// TIA Portal V19 export
DATA_BLOCK "Tacho2_EM02"   // DB3
VERSION : 1.0
// stored: InstanceOfName EM02_Vacio, InstanceOfType FB
"EM02_Vacio"
   // VAR_INPUT
   //    In : "EM02_Input";
   //    VacuumPV : Real := 1000.0;
   //    PumpFbkRun : Bool;
   // END_VAR
   // VAR_OUTPUT
   //    Out : "EM02_Output";
   //    CM_PIC_MV : Real := 100.0;
   //    CM_MotL_Out : Bool := FALSE;
   //    CM_Bk_Out : Bool := FALSE;
   //    TimeoutAlarm : Bool := FALSE;
   //    SensorAlarm : Bool := FALSE;
   //    CMAlarm : Bool := FALSE;
   // END_VAR
   // VAR
   //    State : Int := 1;
   //    ActiveAction : Int := 1;
   //    AlarmLatched : Bool := TRUE;
   //    FaultCode : Int := 4;
   //    TimerReachedSP { S7_SetPoint := 'True'} : TON_TIME;
   //    TimerTimeout { S7_SetPoint := 'True'} : TON_TIME;
   //    TrigStart { S7_SetPoint := 'True'} : R_TRIG;
   //    TrigStop { S7_SetPoint := 'True'} : R_TRIG;
   //    TrigHold { S7_SetPoint := 'True'} : R_TRIG;
   //    TrigAbort { S7_SetPoint := 'True'} : R_TRIG;
   //    TrigReset { S7_SetPoint := 'True'} : R_TRIG;
   //    CM_PIC_Vacuum { S7_SetPoint := 'True'} : "PidL";
   //    CM_MotL { S7_SetPoint := 'True'} : "MotL";
   //    CM_Vlv_Break { S7_SetPoint := 'True'} : "VlvL";
   // END_VAR
BEGIN
   In.Cmds.Start := FALSE;
   In.Cmds.Stop := FALSE;
   In.Cmds.Hold := FALSE;
   In.Cmds.Abort := FALSE;
   In.Cmds.Reset := FALSE;
   In.Cmds.Manual := FALSE;
   In.Cmds.Auto := FALSE;
   In.Cmds.Maintenance := FALSE;
   In.CtrlMode := 0;
   In.VaccumSP := 200.0;
   In.AtmPressure := 980.0;
   In.VaccumValid := TRUE;
   In.VaccumFilter := T#3S;
   In.VaccumTimeout := T#10M;
   In.VaccumSMMV := 0.0;
   Out.Status.ModeMan := FALSE;
   Out.Status.ModeAuto := TRUE;
   Out.Status.ModeMaint := FALSE;
   Out.Status.ModeConflict := FALSE;
   Out.Status.Idle := FALSE;
   Out.Status.Running := TRUE;
   Out.Status.Completed := FALSE;
   Out.Status.Holding := FALSE;
   Out.Status.Held := FALSE;
   Out.Status.Stopping := FALSE;
   Out.Status.Stopped := FALSE;
   Out.Status.Aborting := FALSE;
   Out.Status.Aborted := FALSE;
   Out.Status.Fault := TRUE;
   Out.Status.State := 1;
   Out.Status.FaultCode := 4;
   Out.VacuumActive := TRUE;
   Out.VacuumBroken := FALSE;
   TimerReachedSP.PT := T#0MS;
   TimerReachedSP.IN := FALSE;
   TimerTimeout.PT := T#10M;
   TimerTimeout.IN := TRUE;
   TrigStart.CLK := TRUE;
   TrigStart.Q := FALSE;
   TrigStart.Stat_Bit := TRUE;
   TrigStop.CLK := FALSE;
   TrigStop.Q := FALSE;
   TrigStop.Stat_Bit := FALSE;
   TrigHold.CLK := FALSE;
   TrigHold.Q := FALSE;
   TrigHold.Stat_Bit := FALSE;
   TrigAbort.CLK := FALSE;
   TrigAbort.Q := FALSE;
   TrigAbort.Stat_Bit := FALSE;
   TrigReset.CLK := FALSE;
   TrigReset.Q := FALSE;
   TrigReset.Stat_Bit := FALSE;
   CM_PIC_Vacuum.AutModLi := TRUE;
   CM_PIC_Vacuum.ManModLi := FALSE;
   CM_PIC_Vacuum.LocModLi := FALSE;
   CM_PIC_Vacuum.OosModLi := FALSE;
   CM_PIC_Vacuum.ModLiOp := TRUE;
   CM_PIC_Vacuum.ResetLi := FALSE;
   CM_PIC_Vacuum.SPModLiOp := TRUE;
   CM_PIC_Vacuum.ExtModLi := FALSE;
   CM_PIC_Vacuum.IntModLi := TRUE;
   CM_PIC_Vacuum.PV := 1000.0;
   CM_PIC_Vacuum.PV_Norm.High := 2000.0;
   CM_PIC_Vacuum.PV_Norm.Low := 0.0;
   CM_PIC_Vacuum.MV_Norm.High := 100.0;
   CM_PIC_Vacuum.MV_Norm.Low := 0.0;
   CM_PIC_Vacuum.PV_Scale.High := 2000.0;
   CM_PIC_Vacuum.PV_Scale.Low := 0.0;
   CM_PIC_Vacuum.SPExt := 0.0;
   CM_PIC_Vacuum.SP_HiLim := 2000.0;
   CM_PIC_Vacuum.SP_LoLim := 0.0;
   CM_PIC_Vacuum.MV_HiLim := 100.0;
   CM_PIC_Vacuum.MV_LoLim := 0.0;
   CM_PIC_Vacuum.OosSafeMV := 0.0;
   CM_PIC_Vacuum.PV_unit := 1138;
   CM_PIC_Vacuum.MV_unit := 1342;
   CM_PIC_Vacuum.DataHMI.identName := 'PCV-210';
   CM_PIC_Vacuum.DataHMI.comment := 'Vacio';
   CM_PIC_Vacuum.DataHMI.AutModOp := TRUE;
   CM_PIC_Vacuum.DataHMI.ManModOp := FALSE;
   CM_PIC_Vacuum.DataHMI.LocModOp := FALSE;
   CM_PIC_Vacuum.DataHMI.OosModOp := FALSE;
   CM_PIC_Vacuum.DataHMI.ResetOp := FALSE;
   CM_PIC_Vacuum.DataHMI.MonitorOn := FALSE;
   CM_PIC_Vacuum.DataHMI.ExtModOp := FALSE;
   CM_PIC_Vacuum.DataHMI.IntModOp := FALSE;
   CM_PIC_Vacuum.DataHMI.SpInt := 200.0;
   CM_PIC_Vacuum.DataHMI.Man := 100.0;
   CM_PIC_Vacuum.DataHMI.PermissionLog.AutModOpEn := FALSE;
   CM_PIC_Vacuum.DataHMI.PermissionLog.ManModOpEn := FALSE;
   CM_PIC_Vacuum.DataHMI.PermissionLog.LocModOpEn := FALSE;
   CM_PIC_Vacuum.DataHMI.PermissionLog.OosModOpEn := FALSE;
   CM_PIC_Vacuum.DataHMI.PermissionLog.ResetOpEn := TRUE;
   CM_PIC_Vacuum.DataHMI.PermissionLog.ExtModOpEn := FALSE;
   CM_PIC_Vacuum.DataHMI.PermissionLog.IntModOpEn := FALSE;
   CM_PIC_Vacuum.DataHMI.PermissionLog.Alarms.MsgSupEn := FALSE;
   CM_PIC_Vacuum.DataHMI.PermissionLog.Alarms.HiAlmSupEn := FALSE;
   CM_PIC_Vacuum.DataHMI.PermissionLog.Alarms.HiWrnSupEn := FALSE;
   CM_PIC_Vacuum.DataHMI.PermissionLog.Alarms.LoWrnSupEn := FALSE;
   CM_PIC_Vacuum.DataHMI.PermissionLog.Alarms.LoAlmSupEn := FALSE;
   CM_PIC_Vacuum.DataHMI.Status.OosAct := FALSE;
   CM_PIC_Vacuum.DataHMI.Status.LocAct := FALSE;
   CM_PIC_Vacuum.DataHMI.Status.ManAct := FALSE;
   CM_PIC_Vacuum.DataHMI.Status.AutAct := TRUE;
   CM_PIC_Vacuum.DataHMI.Status.SpExtAct := FALSE;
   CM_PIC_Vacuum.DataHMI.Status.Protection := FALSE;
   CM_PIC_Vacuum.DataHMI.Status.Intlock := TRUE;
   CM_PIC_Vacuum.DataHMI.Status.Permit := TRUE;
   CM_PIC_Vacuum.DataHMI.Status.TrackAct := FALSE;
   CM_PIC_Vacuum.DataHMI.Status.SP := 200.0;
   CM_PIC_Vacuum.DataHMI.Status.PV := 1000.0;
   CM_PIC_Vacuum.DataHMI.Status.ER := -800.0;
   CM_PIC_Vacuum.DataHMI.Status.MV := 100.0;
   CM_PIC_Vacuum.DataHMI.Status.PVOpScale.High := 2000.0;
   CM_PIC_Vacuum.DataHMI.Status.PVOpScale.Low := 0.0;
   CM_PIC_Vacuum.DataHMI.Status.MVOpScale.High := 100.0;
   CM_PIC_Vacuum.DataHMI.Status.MVOpScale.Low := 0.0;
   CM_PIC_Vacuum.DataHMI.Status.SPIntLim.High := 0.0;
   CM_PIC_Vacuum.DataHMI.Status.SPIntLim.Low := 0.0;
   CM_PIC_Vacuum.DataHMI.Status.PV_unit := 1138;
   CM_PIC_Vacuum.DataHMI.Status.MV_unit := 1342;
   CM_PIC_Vacuum.DataHMI.PIDConfig.NegGain := TRUE;
   CM_PIC_Vacuum.DataHMI.PIDConfig.P_Sel := TRUE;
   CM_PIC_Vacuum.DataHMI.PIDConfig.I_Sel := TRUE;
   CM_PIC_Vacuum.DataHMI.PIDConfig.D_Sel := FALSE;
   CM_PIC_Vacuum.DataHMI.PIDConfig.Gain := -2.0;
   CM_PIC_Vacuum.DataHMI.PIDConfig.Ti := 20.0;
   CM_PIC_Vacuum.DataHMI.PIDConfig.Td := 10.0;
   CM_PIC_Vacuum.DataHMI.PIDConfig.DeadBW := 0.0;
   CM_PIC_Vacuum.DataHMI.Alarms.identName := 'PCV-210';
   CM_PIC_Vacuum.DataHMI.Alarms.comment := 'Vacio';
   CM_PIC_Vacuum.DataHMI.Alarms.MsgSupOp := FALSE;
   CM_PIC_Vacuum.DataHMI.Alarms.PVScale.High := 2000.0;
   CM_PIC_Vacuum.DataHMI.Alarms.PVScale.Low := 0.0;
   CM_PIC_Vacuum.DataHMI.Alarms.HiAlmSupOp := FALSE;
   CM_PIC_Vacuum.DataHMI.Alarms.HiWrnSupOp := FALSE;
   CM_PIC_Vacuum.DataHMI.Alarms.LoWrnSupOp := FALSE;
   CM_PIC_Vacuum.DataHMI.Alarms.LoAlmSupOp := FALSE;
   CM_PIC_Vacuum.DataHMI.Alarms.PermissionLog.MsgSupEn := FALSE;
   CM_PIC_Vacuum.DataHMI.Alarms.PermissionLog.HiAlmSupEn := TRUE;
   CM_PIC_Vacuum.DataHMI.Alarms.PermissionLog.HiWrnSupEn := TRUE;
   CM_PIC_Vacuum.DataHMI.Alarms.PermissionLog.LoWrnSupEn := TRUE;
   CM_PIC_Vacuum.DataHMI.Alarms.PermissionLog.LoAlmSupEn := TRUE;
   CM_PIC_Vacuum.DataHMI.Alarms.Status.PV := 1000.0;
   CM_PIC_Vacuum.DataHMI.Alarms.Status.PV_unit := 1138;
   CM_PIC_Vacuum.DataHMI.Alarms.Status.PV_HiAlm := TRUE;
   CM_PIC_Vacuum.DataHMI.Alarms.Status.PV_HiWrn := TRUE;
   CM_PIC_Vacuum.DataHMI.Alarms.Status.PV_LoWrn := FALSE;
   CM_PIC_Vacuum.DataHMI.Alarms.Status.PV_LoAlm := FALSE;
   CM_PIC_Vacuum.DataHMI.Alarms.Status.MsgSup := FALSE;
   CM_PIC_Vacuum.Feature.Startup := TRUE;
   CM_PIC_Vacuum.Feature.MSSOff := TRUE;
   CM_PIC_Vacuum.Feature.FltOff := TRUE;
   CM_PIC_Vacuum.Feature.LocalMod := FALSE;
   CM_PIC_Vacuum.Permission.AutModOpEn := TRUE;
   CM_PIC_Vacuum.Permission.ManModOpEn := TRUE;
   CM_PIC_Vacuum.Permission.LocModOpEn := FALSE;
   CM_PIC_Vacuum.Permission.OosModOpEn := FALSE;
   CM_PIC_Vacuum.Permission.ResetOpEn := TRUE;
   CM_PIC_Vacuum.Permission.ExtModOpEn := FALSE;
   CM_PIC_Vacuum.Permission.IntModOpEn := TRUE;
   CM_PIC_Vacuum.Permission.Alarms.MsgSupEn := TRUE;
   CM_PIC_Vacuum.Permission.Alarms.HiAlmSupEn := TRUE;
   CM_PIC_Vacuum.Permission.Alarms.HiWrnSupEn := TRUE;
   CM_PIC_Vacuum.Permission.Alarms.LoWrnSupEn := TRUE;
   CM_PIC_Vacuum.Permission.Alarms.LoAlmSupEn := TRUE;
   CM_PIC_Vacuum.MSS := TRUE;
   CM_PIC_Vacuum.Trip := FALSE;
   CM_PIC_Vacuum.Permit := TRUE;
   CM_PIC_Vacuum.Intlock := TRUE;
   CM_PIC_Vacuum.Protect := TRUE;
   CM_PIC_Vacuum.TrackOn := FALSE;
   CM_PIC_Vacuum.Rbk := 0.0;
   CM_PIC_Vacuum.RbkHiTol := 3.0;
   CM_PIC_Vacuum.RbkLoTol := 3.0;
   CM_PIC_Vacuum.RbkMonTime := T#3S;
   CM_PIC_Vacuum.TrackVal := 0.0;
   CM_PIC_Vacuum.RunUpCyc := 3;
   CM_PIC_Vacuum.DisV := 0.0;
   CM_PIC_Vacuum.HiAlm := 95.0;
   CM_PIC_Vacuum.HiWrn := 90.0;
   CM_PIC_Vacuum.LoWrn := 10.0;
   CM_PIC_Vacuum.LoAlm := 5.0;
   CM_PIC_Vacuum.Hyst := 5.0;
   CM_PIC_Vacuum.AutAct := TRUE;
   CM_PIC_Vacuum.ManAct := FALSE;
   CM_PIC_Vacuum.LocAct := FALSE;
   CM_PIC_Vacuum.OosAct := FALSE;
   CM_PIC_Vacuum.MsgSup := TRUE;
   CM_PIC_Vacuum.AlarmError := FALSE;
   CM_PIC_Vacuum.MV := 100.0;
   CM_PIC_Vacuum.SPExtAct := FALSE;
   CM_PIC_Vacuum.SP := 200.0;
   CM_PIC_Vacuum.ER := -800.0;
   CM_PIC_Vacuum.PVH_Alm := TRUE;
   CM_PIC_Vacuum.PVH_Wrn := TRUE;
   CM_PIC_Vacuum.PVL_Wrn := FALSE;
   CM_PIC_Vacuum.PVL_Alm := FALSE;
   CM_PIC_Vacuum.controller.COM_RST := FALSE;
   CM_PIC_Vacuum.controller.MAN_ON := FALSE;
   CM_PIC_Vacuum.controller.PVPER_ON := FALSE;
   CM_PIC_Vacuum.controller.P_SEL := TRUE;
   CM_PIC_Vacuum.controller.I_SEL := TRUE;
   CM_PIC_Vacuum.controller.INT_HOLD := FALSE;
   CM_PIC_Vacuum.controller.I_ITL_ON := FALSE;
   CM_PIC_Vacuum.controller.D_SEL := FALSE;
   CM_PIC_Vacuum.controller.CYCLE := T#1S;
   CM_PIC_Vacuum.controller.SP_INT := 10.0;
   CM_PIC_Vacuum.controller.PV_IN := 50.0;
   CM_PIC_Vacuum.controller.PV_PER := 16#0000;
   CM_PIC_Vacuum.controller.MAN := 100.0;
   CM_PIC_Vacuum.controller.GAIN := -2.0;
   CM_PIC_Vacuum.controller.TI := T#20S;
   CM_PIC_Vacuum.controller.TD := T#10S;
   CM_PIC_Vacuum.controller.TM_LAG := T#2S;
   CM_PIC_Vacuum.controller.DEADB_W := 0.0;
   CM_PIC_Vacuum.controller.LMN_HLM := 100.0;
   CM_PIC_Vacuum.controller.LMN_LLM := 0.0;
   CM_PIC_Vacuum.controller.PV_FAC := 1.0;
   CM_PIC_Vacuum.controller.PV_OFF := 0.0;
   CM_PIC_Vacuum.controller.LMN_FAC := 1.0;
   CM_PIC_Vacuum.controller.LMN_OFF := 0.0;
   CM_PIC_Vacuum.controller.I_ITLVAL := 0.0;
   CM_PIC_Vacuum.controller.DISV := 0.0;
   CM_PIC_Vacuum.controller.LMN := 100.0;
   CM_PIC_Vacuum.controller.LMN_PER := 16#6C00;
   CM_PIC_Vacuum.controller.QLMN_HLM := TRUE;
   CM_PIC_Vacuum.controller.QLMN_LLM := FALSE;
   CM_PIC_Vacuum.controller.LMN_P := 80.0;
   CM_PIC_Vacuum.controller.LMN_I := 80.0;
   CM_PIC_Vacuum.controller.LMN_D := 0.0;
   CM_PIC_Vacuum.controller.PV := 50.0;
   CM_PIC_Vacuum.controller.ER := -40.0;
   CM_PIC_Vacuum.controller.sInvAlt := 80.0;
   CM_PIC_Vacuum.controller.sIanteilAlt := 80.0;
   CM_PIC_Vacuum.controller.sRestInt := 0.0;
   CM_PIC_Vacuum.controller.sRestDif := 0.0;
   CM_PIC_Vacuum.controller.sRueck := 80.0;
   CM_PIC_Vacuum.controller.sLmn := 100.0;
   CM_PIC_Vacuum.controller.sbArwHLmOn := TRUE;
   CM_PIC_Vacuum.controller.sbArwLLmOn := FALSE;
   CM_PIC_Vacuum.controller.sbILimOn := TRUE;
   CM_PIC_Vacuum.ModSelInt := 2;
   CM_PIC_Vacuum.stRestart := FALSE;
   CM_PIC_Vacuum.ResetLiLogic := FALSE;
   CM_PIC_Vacuum.ResetResult := FALSE;
   CM_PIC_Vacuum.stResetLiLogic := FALSE;
   CM_PIC_Vacuum.stMonErr := FALSE;
   CM_PIC_Vacuum.stTripErr := FALSE;
   CM_PIC_Vacuum.stProtErr := FALSE;
   CM_PIC_Vacuum.stMSS := FALSE;
   CM_PIC_Vacuum.stProt := FALSE;
   CM_PIC_Vacuum.stTrip := FALSE;
   CM_PIC_Vacuum.stLockFault := FALSE;
   CM_PIC_Vacuum.stRun := FALSE;
   CM_PIC_Vacuum.stExtMod := FALSE;
   CM_PIC_Vacuum.stAutoLogic := FALSE;
   CM_PIC_Vacuum.RuntimeMem := 16#0000_0EAA_9B49_C0F5;
   CM_PIC_Vacuum.RuntimeS := 0.999710415986597;
   CM_PIC_Vacuum.PVMon.Feature.Startup := TRUE;
   CM_PIC_Vacuum.PVMon.Enable := TRUE;
   CM_PIC_Vacuum.PVMon.Permission.MsgSupEn := TRUE;
   CM_PIC_Vacuum.PVMon.Permission.HiAlmSupEn := TRUE;
   CM_PIC_Vacuum.PVMon.Permission.HiWrnSupEn := TRUE;
   CM_PIC_Vacuum.PVMon.Permission.LoWrnSupEn := TRUE;
   CM_PIC_Vacuum.PVMon.Permission.LoAlmSupEn := TRUE;
   CM_PIC_Vacuum.PVMon.DataHMI.identName := 'PCV-210';
   CM_PIC_Vacuum.PVMon.DataHMI.comment := 'Vacio';
   CM_PIC_Vacuum.PVMon.DataHMI.MsgSupOp := FALSE;
   CM_PIC_Vacuum.PVMon.DataHMI.PVScale.High := 2000.0;
   CM_PIC_Vacuum.PVMon.DataHMI.PVScale.Low := 0.0;
   CM_PIC_Vacuum.PVMon.DataHMI.HiAlmSupOp := FALSE;
   CM_PIC_Vacuum.PVMon.DataHMI.HiWrnSupOp := FALSE;
   CM_PIC_Vacuum.PVMon.DataHMI.LoWrnSupOp := FALSE;
   CM_PIC_Vacuum.PVMon.DataHMI.LoAlmSupOp := FALSE;
   CM_PIC_Vacuum.PVMon.DataHMI.PermissionLog.MsgSupEn := FALSE;
   CM_PIC_Vacuum.PVMon.DataHMI.PermissionLog.HiAlmSupEn := TRUE;
   CM_PIC_Vacuum.PVMon.DataHMI.PermissionLog.HiWrnSupEn := TRUE;
   CM_PIC_Vacuum.PVMon.DataHMI.PermissionLog.LoWrnSupEn := TRUE;
   CM_PIC_Vacuum.PVMon.DataHMI.PermissionLog.LoAlmSupEn := TRUE;
   CM_PIC_Vacuum.PVMon.DataHMI.Status.PV := 1000.0;
   CM_PIC_Vacuum.PVMon.DataHMI.Status.PV_unit := 1138;
   CM_PIC_Vacuum.PVMon.DataHMI.Status.PV_HiAlm := TRUE;
   CM_PIC_Vacuum.PVMon.DataHMI.Status.PV_HiWrn := TRUE;
   CM_PIC_Vacuum.PVMon.DataHMI.Status.PV_LoWrn := FALSE;
   CM_PIC_Vacuum.PVMon.DataHMI.Status.PV_LoAlm := FALSE;
   CM_PIC_Vacuum.PVMon.DataHMI.Status.MsgSup := FALSE;
   CM_PIC_Vacuum.PVMon.RunUpCyc := 3;
   CM_PIC_Vacuum.PVMon.PV := 1000.0;
   CM_PIC_Vacuum.PVMon.HiAlm := 95.0;
   CM_PIC_Vacuum.PVMon.HiWrn := 90.0;
   CM_PIC_Vacuum.PVMon.LoWrn := 10.0;
   CM_PIC_Vacuum.PVMon.LoAlm := 5.0;
   CM_PIC_Vacuum.PVMon.Hyst := 5.0;
   CM_PIC_Vacuum.PVMon.PV_unit := 1138;
   CM_PIC_Vacuum.PVMon.MsgErr := FALSE;
   CM_PIC_Vacuum.PVMon.MsgSup := TRUE;
   CM_PIC_Vacuum.PVMon.PVH_Alm := TRUE;
   CM_PIC_Vacuum.PVMon.PVH_Wrn := TRUE;
   CM_PIC_Vacuum.PVMon.PVL_Wrn := FALSE;
   CM_PIC_Vacuum.PVMon.PVL_Alm := FALSE;
   CM_PIC_Vacuum.PVMon.stRestart := FALSE;
   CM_PIC_Vacuum.PVMon.RunUpCounter := 0;
   CM_PIC_Vacuum.PVMon.pSIG1 := TRUE;
   CM_PIC_Vacuum.PVMon.pSIG2 := TRUE;
   CM_PIC_Vacuum.PVMon.pSIG3 := FALSE;
   CM_PIC_Vacuum.PVMon.pSIG4 := FALSE;
   CM_PIC_Vacuum.PVMon.pAlarm := TRUE;
   CM_PIC_Vacuum.RunUpCounter := 0;
   CM_PIC_Vacuum.pAlarm := TRUE;
   CM_PIC_Vacuum.stMSSErr := FALSE;
   CM_PIC_Vacuum.SPMod := FALSE;
   CM_PIC_Vacuum.SPSelInt := 1;
   CM_PIC_Vacuum.stErr := FALSE;
   CM_PIC_Vacuum.stDivErr := FALSE;
   CM_PIC_Vacuum.stNegGain := TRUE;
   CM_PIC_Vacuum.stGain := -2.0;
   CM_PIC_Vacuum.stTi := 0.0;
   CM_PIC_Vacuum.stTd := 0.0;
   CM_PIC_Vacuum.stPIDConfig.NegGain := TRUE;
   CM_PIC_Vacuum.stPIDConfig.P_Sel := TRUE;
   CM_PIC_Vacuum.stPIDConfig.I_Sel := TRUE;
   CM_PIC_Vacuum.stPIDConfig.D_Sel := FALSE;
   CM_PIC_Vacuum.stPIDConfig.Gain := -2.0;
   CM_PIC_Vacuum.stPIDConfig.Ti := 20.0;
   CM_PIC_Vacuum.stPIDConfig.Td := 10.0;
   CM_PIC_Vacuum.stPIDConfig.DeadBW := 0.0;
   CM_PIC_Vacuum.RbkMonitorTimer.PT := T#0MS;
   CM_PIC_Vacuum.RbkMonitorTimer.IN := FALSE;
   CM_MotL.SampleT := 1.0;
   CM_MotL.AutModLi := TRUE;
   CM_MotL.ManModLi := FALSE;
   CM_MotL.LocModLi := FALSE;
   CM_MotL.OosModLi := FALSE;
   CM_MotL.ModLiOp := TRUE;
   CM_MotL.ResetLi := FALSE;
   CM_MotL.DataHMI.identName := 'M-102';
   CM_MotL.DataHMI.comment := 'Bba Vacio';
   CM_MotL.DataHMI.AutModOp := TRUE;
   CM_MotL.DataHMI.ManModOp := FALSE;
   CM_MotL.DataHMI.LocModOp := FALSE;
   CM_MotL.DataHMI.OosModOp := FALSE;
   CM_MotL.DataHMI.StartOp := FALSE;
   CM_MotL.DataHMI.StopOp := FALSE;
   CM_MotL.DataHMI.ResetOp := FALSE;
   CM_MotL.DataHMI.MonitorOn := FALSE;
   CM_MotL.DataHMI.PermissionLog.AutModOpEn := FALSE;
   CM_MotL.DataHMI.PermissionLog.ManModOpEn := FALSE;
   CM_MotL.DataHMI.PermissionLog.LocModOpEn := FALSE;
   CM_MotL.DataHMI.PermissionLog.OosModOpEn := FALSE;
   CM_MotL.DataHMI.PermissionLog.ResetOpEn := TRUE;
   CM_MotL.DataHMI.PermissionLog.StartOpEn := FALSE;
   CM_MotL.DataHMI.PermissionLog.StopOpEn := FALSE;
   CM_MotL.DataHMI.Status.OosAct := FALSE;
   CM_MotL.DataHMI.Status.LocAct := FALSE;
   CM_MotL.DataHMI.Status.ManAct := FALSE;
   CM_MotL.DataHMI.Status.AutAct := TRUE;
   CM_MotL.DataHMI.Status.CmdOnOff := TRUE;
   CM_MotL.DataHMI.Status.Run := TRUE;
   CM_MotL.DataHMI.Status.Stop := FALSE;
   CM_MotL.DataHMI.Status.MonErr := FALSE;
   CM_MotL.DataHMI.Status.Trip := FALSE;
   CM_MotL.DataHMI.Status.Protection := FALSE;
   CM_MotL.DataHMI.Status.Intlock := TRUE;
   CM_MotL.DataHMI.Status.Permit := TRUE;
   CM_MotL.DataHMI.MonitorTime := 3.0;
   CM_MotL.Feature.Startup := TRUE;
   CM_MotL.Feature.MSSOff := TRUE;
   CM_MotL.Feature.FltOff := TRUE;
   CM_MotL.Feature.LocalMod := FALSE;
   CM_MotL.Permission.AutModOpEn := TRUE;
   CM_MotL.Permission.ManModOpEn := TRUE;
   CM_MotL.Permission.LocModOpEn := FALSE;
   CM_MotL.Permission.OosModOpEn := FALSE;
   CM_MotL.Permission.ResetOpEn := TRUE;
   CM_MotL.Permission.StartOpEn := TRUE;
   CM_MotL.Permission.StopOpEn := TRUE;
   CM_MotL.MSS := TRUE;
   CM_MotL.Trip := FALSE;
   CM_MotL.Permit := TRUE;
   CM_MotL.Intlock := TRUE;
   CM_MotL.Protect := TRUE;
   CM_MotL.StartAut := TRUE;
   CM_MotL.StopAut := FALSE;
   CM_MotL.StartLoc := FALSE;
   CM_MotL.StopLoc := FALSE;
   CM_MotL.LockOn := FALSE;
   CM_MotL.FbkRun := FALSE;
   CM_MotL.RunUpCyc := 3;
   CM_MotL.Start := TRUE;
   CM_MotL.AutAct := TRUE;
   CM_MotL.ManAct := FALSE;
   CM_MotL.LocAct := FALSE;
   CM_MotL.OosAct := FALSE;
   CM_MotL.Run := TRUE;
   CM_MotL.Stop := FALSE;
   CM_MotL.MsgSup := FALSE;
   CM_MotL.AlarmError := FALSE;
   CM_MotL.ModSelInt := 2;
   CM_MotL.stRestart := FALSE;
   CM_MotL.ResetLiLogic := FALSE;
   CM_MotL.ResetResult := FALSE;
   CM_MotL.stResetLiLogic := FALSE;
   CM_MotL.stMonErr := FALSE;
   CM_MotL.stTripErr := FALSE;
   CM_MotL.stProtErr := FALSE;
   CM_MotL.stMSS := FALSE;
   CM_MotL.stProt := FALSE;
   CM_MotL.stTrip := FALSE;
   CM_MotL.stLockFault := FALSE;
   CM_MotL.stRun := TRUE;
   CM_MotL.stCmdOnOff := TRUE;
   CM_MotL.stAutoLogic := TRUE;
   CM_MotL.stbCmdOnOff := TRUE;
   CM_MotL.stActiveTime := 0.0;
   CM_MotL.RunUpCounter := 0;
   CM_MotL.pAlarm := TRUE;
   CM_MotL.stMSSErr := FALSE;
   CM_Vlv_Break.SampleT := 1.0;
   CM_Vlv_Break.AutModLi := TRUE;
   CM_Vlv_Break.ManModLi := FALSE;
   CM_Vlv_Break.LocModLi := FALSE;
   CM_Vlv_Break.OosModLi := FALSE;
   CM_Vlv_Break.ModLiOp := TRUE;
   CM_Vlv_Break.ResetLi := FALSE;
   CM_Vlv_Break.DataHMI.identName := 'PSV-103';
   CM_Vlv_Break.DataHMI.comment := 'Rompevacio';
   CM_Vlv_Break.DataHMI.AutModOp := TRUE;
   CM_Vlv_Break.DataHMI.ManModOp := FALSE;
   CM_Vlv_Break.DataHMI.LocModOp := FALSE;
   CM_Vlv_Break.DataHMI.OosModOp := FALSE;
   CM_Vlv_Break.DataHMI.OpenOp := FALSE;
   CM_Vlv_Break.DataHMI.CloseOp := FALSE;
   CM_Vlv_Break.DataHMI.ResetOp := FALSE;
   CM_Vlv_Break.DataHMI.MonitorOn := FALSE;
   CM_Vlv_Break.DataHMI.PermissionLog.AutModOpEn := FALSE;
   CM_Vlv_Break.DataHMI.PermissionLog.ManModOpEn := FALSE;
   CM_Vlv_Break.DataHMI.PermissionLog.LocModOpEn := FALSE;
   CM_Vlv_Break.DataHMI.PermissionLog.OosModOpEn := FALSE;
   CM_Vlv_Break.DataHMI.PermissionLog.ResetOpEn := TRUE;
   CM_Vlv_Break.DataHMI.PermissionLog.OpenOpEn := FALSE;
   CM_Vlv_Break.DataHMI.PermissionLog.CloseOpEn := FALSE;
   CM_Vlv_Break.DataHMI.Status.OosAct := FALSE;
   CM_Vlv_Break.DataHMI.Status.LocAct := FALSE;
   CM_Vlv_Break.DataHMI.Status.ManAct := FALSE;
   CM_Vlv_Break.DataHMI.Status.AutAct := TRUE;
   CM_Vlv_Break.DataHMI.Status.Cmd := FALSE;
   CM_Vlv_Break.DataHMI.Status.Opened := FALSE;
   CM_Vlv_Break.DataHMI.Status.Closed := TRUE;
   CM_Vlv_Break.DataHMI.Status.MonErr := FALSE;
   CM_Vlv_Break.DataHMI.Status.Trip := FALSE;
   CM_Vlv_Break.DataHMI.Status.Protection := FALSE;
   CM_Vlv_Break.DataHMI.Status.Intlock := FALSE;
   CM_Vlv_Break.DataHMI.Status.Permit := FALSE;
   CM_Vlv_Break.DataHMI.MonitorTime := 3.0;
   CM_Vlv_Break.Feature.Startup := TRUE;
   CM_Vlv_Break.Feature.MSSOff := TRUE;
   CM_Vlv_Break.Feature.FltOff := TRUE;
   CM_Vlv_Break.Feature.LocalMod := FALSE;
   CM_Vlv_Break.Permission.AutModOpEn := TRUE;
   CM_Vlv_Break.Permission.ManModOpEn := TRUE;
   CM_Vlv_Break.Permission.LocModOpEn := FALSE;
   CM_Vlv_Break.Permission.OosModOpEn := FALSE;
   CM_Vlv_Break.Permission.ResetOpEn := TRUE;
   CM_Vlv_Break.Permission.OpenOpEn := TRUE;
   CM_Vlv_Break.Permission.CloseOpEn := TRUE;
   CM_Vlv_Break.MSS := TRUE;
   CM_Vlv_Break.Trip := FALSE;
   CM_Vlv_Break.Permit := FALSE;
   CM_Vlv_Break.Intlock := FALSE;
   CM_Vlv_Break.Protect := TRUE;
   CM_Vlv_Break.OpenAut := FALSE;
   CM_Vlv_Break.CloseAut := TRUE;
   CM_Vlv_Break.OpenLoc := FALSE;
   CM_Vlv_Break.CloseLoc := FALSE;
   CM_Vlv_Break.LockOn := FALSE;
   CM_Vlv_Break.FbkOpen := FALSE;
   CM_Vlv_Break.FbkClose := FALSE;
   CM_Vlv_Break.SafePos := FALSE;
   CM_Vlv_Break.RunUpCyc := 3;
   CM_Vlv_Break.AutAct := TRUE;
   CM_Vlv_Break.ManAct := FALSE;
   CM_Vlv_Break.LocAct := FALSE;
   CM_Vlv_Break.OosAct := FALSE;
   CM_Vlv_Break.Opened := FALSE;
   CM_Vlv_Break.Closed := TRUE;
   CM_Vlv_Break.MsgSup := FALSE;
   CM_Vlv_Break.AlarmError := FALSE;
   CM_Vlv_Break.cmd := FALSE;
   CM_Vlv_Break.ModSelInt := 2;
   CM_Vlv_Break.stRestart := FALSE;
   CM_Vlv_Break.ResetLiLogic := FALSE;
   CM_Vlv_Break.ResetResult := FALSE;
   CM_Vlv_Break.stResetLiLogic := FALSE;
   CM_Vlv_Break.stMonErr := FALSE;
   CM_Vlv_Break.stTripErr := FALSE;
   CM_Vlv_Break.stProtErr := FALSE;
   CM_Vlv_Break.stMSS := FALSE;
   CM_Vlv_Break.stProt := FALSE;
   CM_Vlv_Break.stTrip := FALSE;
   CM_Vlv_Break.stLockFault := TRUE;
   CM_Vlv_Break.stPosition := FALSE;
   CM_Vlv_Break.stCmd := FALSE;
   CM_Vlv_Break.stAutoLogic := FALSE;
   CM_Vlv_Break.stbCmd := FALSE;
   CM_Vlv_Break.stActiveTime := 0.0;
   CM_Vlv_Break.RunUpCounter := 0;
   CM_Vlv_Break.pAlarm := TRUE;
   CM_Vlv_Break.stMSSErr := FALSE;
END_DATA_BLOCK
